(* Logix 5000 project; controller TFF vendor 1 type 14 code 107 rev 34.11; software revision 34.03; part 24 of 36 *)
(* tags used below, declared in another part *)
   Address : DINT;   // Temp Address
   Address2 : DINT;   // Temp Address
   Index : DINT;   // Index
   ONS_PID02 : BOOL;
   PCV001_PID_Settings : INT;
   AnalogOutput : AnalogOutput[25];   // Analog Output Array
   AnalogPoint : AnalogInput[50];   // Analog Input Array
   ControlLoop : ControlLoop[20];   // Control Loop Array
   ControlLoop_FeedPump : ALIAS FOR ControlLoop[1];   // Feed Pump Control Loop
   ControlLoop_PCV001 : ALIAS FOR ControlLoop[3];   // PCV001 Control Loop
   ControlLoop_PCV001_5ms : ALIAS FOR ControlLoop[4];   // PCV001 Control Loop
   ControlLoop_PCV001_CV : REAL;   // Control Value
   ControlLoop_PCV001_RAMP_OUT : REAL;   // Ramp Output
   ControlLoop_PCV101 : ALIAS FOR ControlLoop[5];   // PCV101 Control Loop
   ControlLoop_PCV101_5ms : ALIAS FOR ControlLoop[6];   // PCV101 Control Loop
   ControlLoop_PCV101_RAMP_OUT : REAL;   // Ramp Output
   PCV001_Control : PCV_Control;   // PCV001 Control UDT
   PCV101 : ALIAS FOR AnalogPoint[4];   // Filtrate Pressure Control Valve Position
   PCV101_Control : PCV_Control;   // PCV101 Control UDT
   PumpRunStatus : DINT;   // Pumps Run Status (1 = At least one pump running , 0 = no pump running)
   SysControl : SysControl;   // General system status and command
(* Process, continued *)

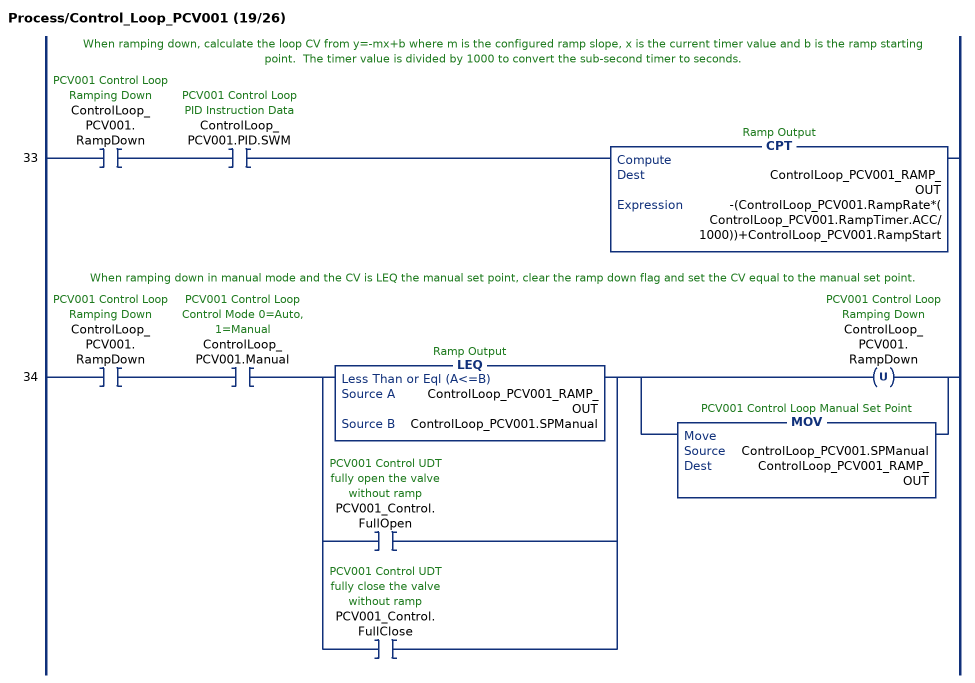
   [picture p213: Process/Control_Loop_PCV001 rungs 33-34]
   // When ramping down, calculate the loop CV from y=-mx+b where m is the configured ramp slope, x is the current timer value and b is the ramp starting point.  The timer value is divided by 1000 to convert the sub-second timer to seconds.
   33: XIC(ControlLoop_PCV001.RampDown)XIC(ControlLoop_PCV001.PID.SWM)CPT(ControlLoop_PCV001_RAMP_OUT,-(ControlLoop_PCV001.RampRate*(ControlLoop_PCV001.RampTimer.ACC/1000))+ControlLoop_PCV001.RampStart);
   // When ramping down in manual mode and the CV is LEQ the manual set point, clear the ramp down flag and set the CV equal to the manual set point.
   34: XIC(ControlLoop_PCV001.RampDown)XIC(ControlLoop_PCV001.Manual)[LEQ(ControlLoop_PCV001_RAMP_OUT,ControlLoop_PCV001.SPManual) ,XIC(PCV001_Control.FullOpen) ,XIC(PCV001_Control.FullClose) ][OTU(ControlLoop_PCV001.RampDown) ,MOV(ControlLoop_PCV001.SPManual,ControlLoop_PCV001_RAMP_OUT) ];
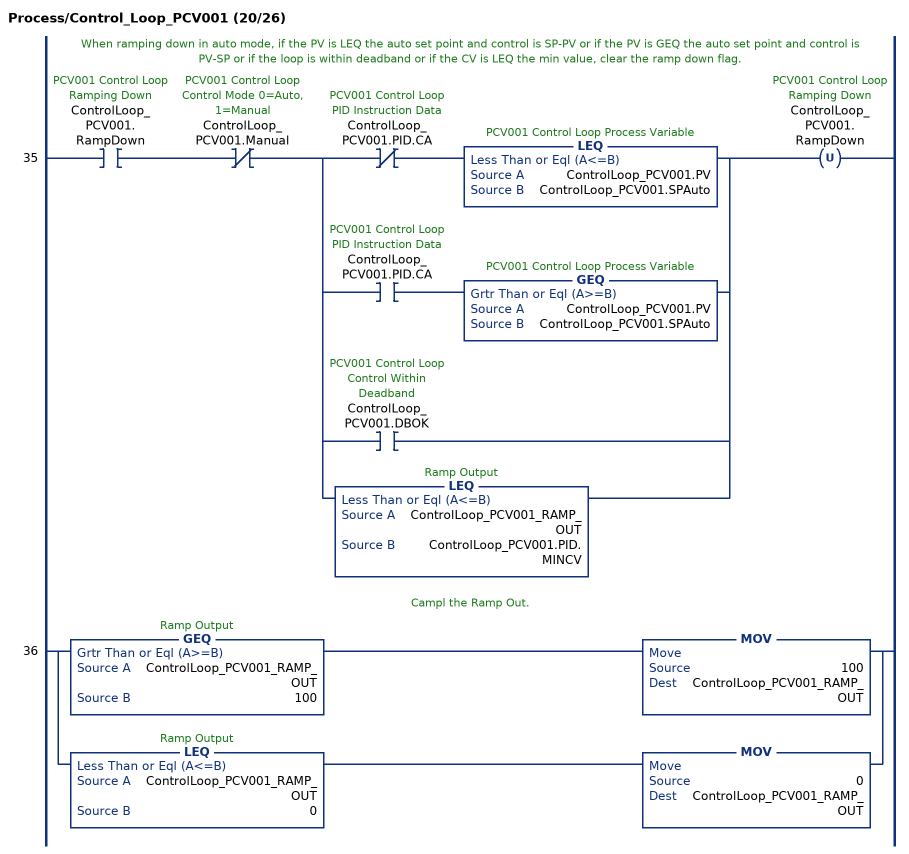
   // When ramping down in auto mode, if the PV is LEQ the auto set point and control is SP-PV or if the PV is GEQ the auto set point and control is PV-SP or if the loop is within deadband or if the CV is LEQ the min value, clear the ramp down flag.
   35: XIC(ControlLoop_PCV001.RampDown)XIO(ControlLoop_PCV001.Manual)[XIO(ControlLoop_PCV001.PID.CA) LEQ(ControlLoop_PCV001.PV,ControlLoop_PCV001.SPAuto) ,XIC(ControlLoop_PCV001.PID.CA) GEQ(ControlLoop_PCV001.PV,ControlLoop_PCV001.SPAuto) ,XIC(ControlLoop_PCV001.DBOK) ,LEQ(ControlLoop_PCV001_RAMP_OUT,ControlLoop_PCV001.PID.MINCV) ]OTU(ControlLoop_PCV001.RampDown);
   // Campl the Ramp Out.
   36: [GEQ(ControlLoop_PCV001_RAMP_OUT,100) MOV(100,ControlLoop_PCV001_RAMP_OUT) ,LEQ(ControlLoop_PCV001_RAMP_OUT,0) MOV(0,ControlLoop_PCV001_RAMP_OUT) ];
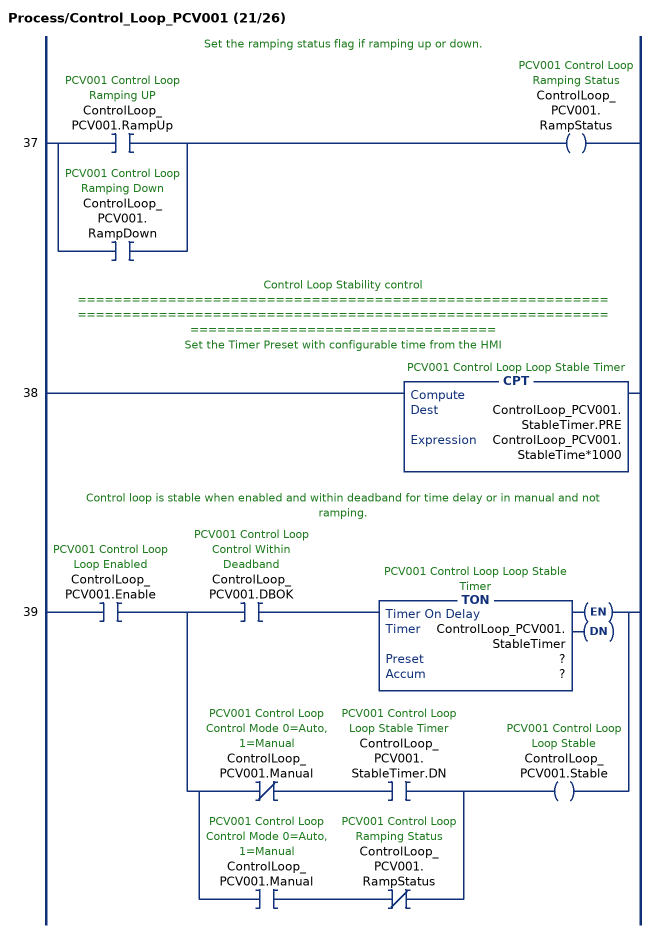
   // Set the ramping status flag if ramping up or down.
   37: [XIC(ControlLoop_PCV001.RampUp) ,XIC(ControlLoop_PCV001.RampDown) ]OTE(ControlLoop_PCV001.RampStatus);
   // Control Loop Stability control
   // ========================================================================================================================================================
   // Set the Timer Preset with configurable time from the HMI
   38: CPT(ControlLoop_PCV001.StableTimer.PRE,ControlLoop_PCV001.StableTime*1000);
   // Control loop is stable when enabled and within deadband for time delay or in manual and not ramping.
   39: XIC(ControlLoop_PCV001.Enable)[XIC(ControlLoop_PCV001.DBOK) TON(ControlLoop_PCV001.StableTimer,?,?) ,[XIO(ControlLoop_PCV001.Manual) XIC(ControlLoop_PCV001.StableTimer.DN) ,XIC(ControlLoop_PCV001.Manual) XIO(ControlLoop_PCV001.RampStatus) ] OTE(ControlLoop_PCV001.Stable) ];
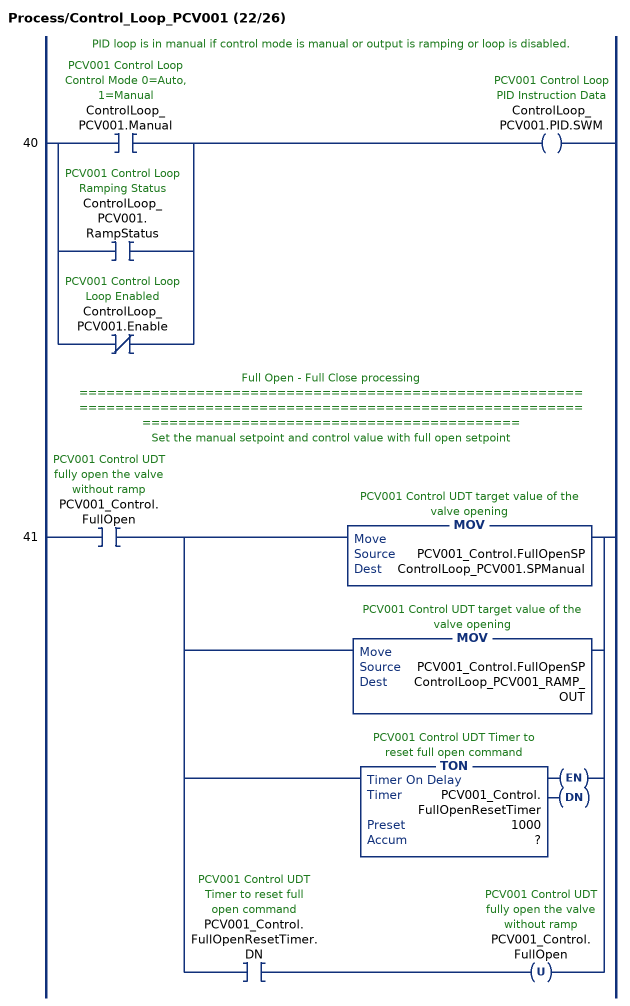
   // PID loop is in manual if control mode is manual or output is ramping or loop is disabled.
   40: [XIC(ControlLoop_PCV001.Manual) ,XIC(ControlLoop_PCV001.RampStatus) ,XIO(ControlLoop_PCV001.Enable) ]OTE(ControlLoop_PCV001.PID.SWM);
   // Full Open - Full Close processing
   // ==========================================================================================================================================================
   // Set the manual setpoint and control value with full open setpoint
   41: XIC(PCV001_Control.FullOpen)[MOV(PCV001_Control.FullOpenSP,ControlLoop_PCV001.SPManual) ,MOV(PCV001_Control.FullOpenSP,ControlLoop_PCV001_RAMP_OUT) ,TON(PCV001_Control.FullOpenResetTimer,?,?) ,XIC(PCV001_Control.FullOpenResetTimer.DN) OTU(PCV001_Control.FullOpen) ];
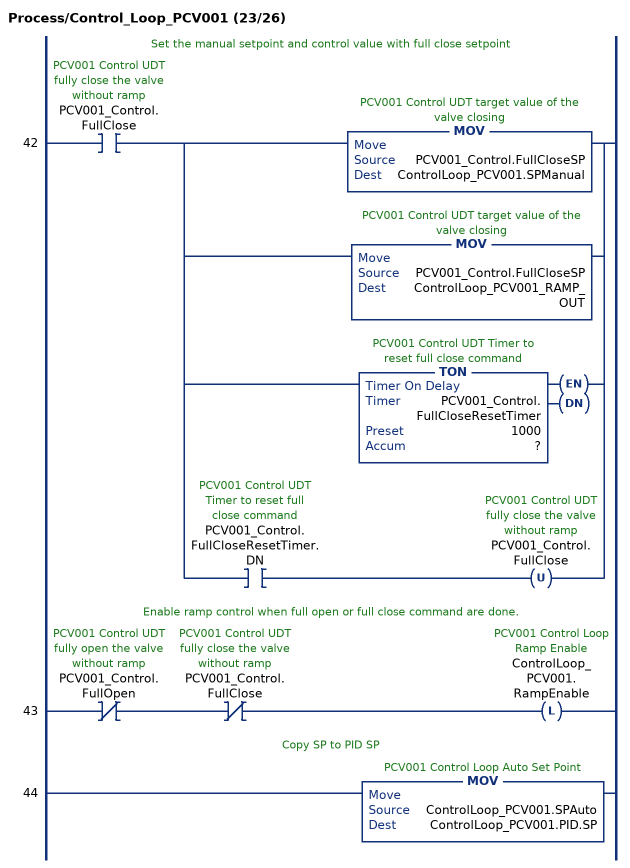
   // Set the manual setpoint and control value with full close setpoint
   42: XIC(PCV001_Control.FullClose)[MOV(PCV001_Control.FullCloseSP,ControlLoop_PCV001.SPManual) ,MOV(PCV001_Control.FullCloseSP,ControlLoop_PCV001_RAMP_OUT) ,TON(PCV001_Control.FullCloseResetTimer,?,?) ,XIC(PCV001_Control.FullCloseResetTimer.DN) OTU(PCV001_Control.FullClose) ];
   // Enable ramp control when full open or full close command are done.
   43: XIO(PCV001_Control.FullOpen)XIO(PCV001_Control.FullClose)OTL(ControlLoop_PCV001.RampEnable);
   // Copy SP to PID SP
   44: MOV(ControlLoop_PCV001.SPAuto,ControlLoop_PCV001.PID.SP);
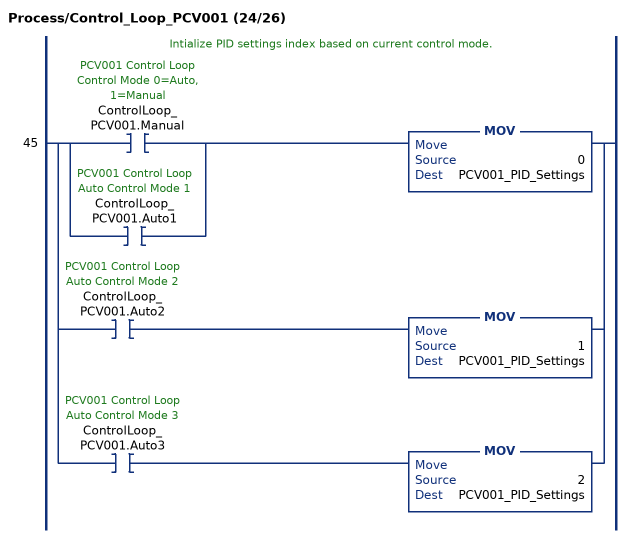
   // Intialize PID settings index based on current control mode.
   45: [[XIC(ControlLoop_PCV001.Manual) ,XIC(ControlLoop_PCV001.Auto1) ] MOV(0,PCV001_PID_Settings) ,XIC(ControlLoop_PCV001.Auto2) MOV(1,PCV001_PID_Settings) ,XIC(ControlLoop_PCV001.Auto3) MOV(2,PCV001_PID_Settings) ];
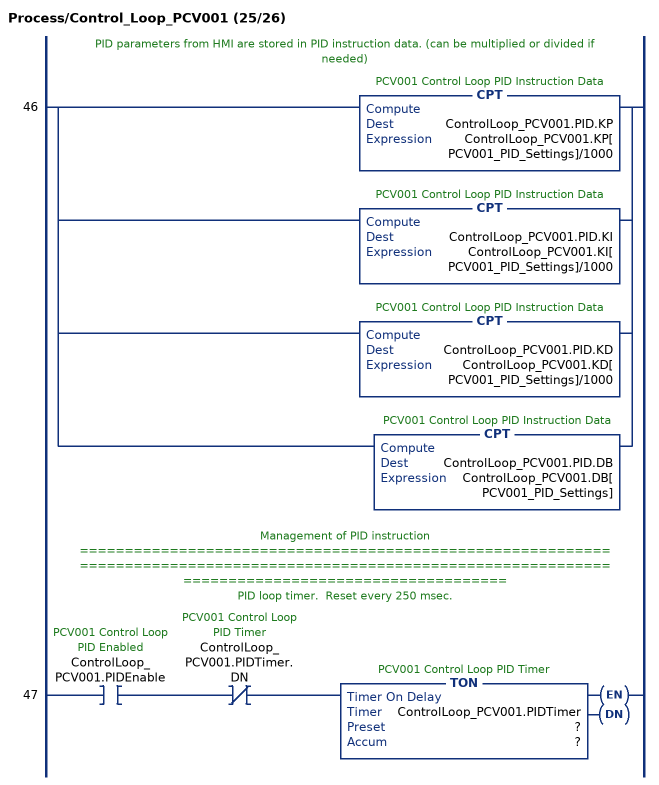
   // PID parameters from HMI are stored in PID instruction data. (can be multiplied or divided if needed)
   46: [CPT(ControlLoop_PCV001.PID.KP,ControlLoop_PCV001.KP[PCV001_PID_Settings]/1000) ,CPT(ControlLoop_PCV001.PID.KI,ControlLoop_PCV001.KI[PCV001_PID_Settings]/1000) ,CPT(ControlLoop_PCV001.PID.KD,ControlLoop_PCV001.KD[PCV001_PID_Settings]/1000) ,CPT(ControlLoop_PCV001.PID.DB,ControlLoop_PCV001.DB[PCV001_PID_Settings]) ];
   // Management of PID instruction
   // ==========================================================================================================================================================
   // PID loop timer.  Reset every 250 msec.
   47: XIC(ControlLoop_PCV001.PIDEnable)XIO(ControlLoop_PCV001.PIDTimer.DN)TON(ControlLoop_PCV001.PIDTimer,?,?);
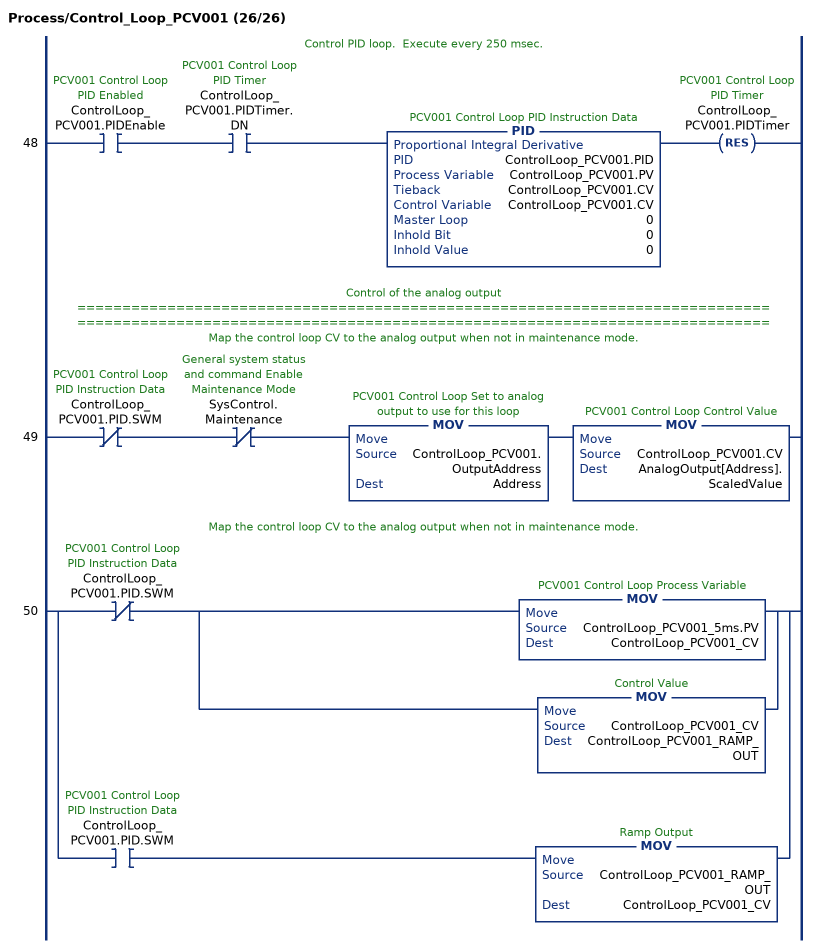
   // Control PID loop.  Execute every 250 msec.
   48: XIC(ControlLoop_PCV001.PIDEnable)XIC(ControlLoop_PCV001.PIDTimer.DN)PID(ControlLoop_PCV001.PID,ControlLoop_PCV001.PV,ControlLoop_PCV001.CV,ControlLoop_PCV001.CV,0,0,0)RES(ControlLoop_PCV001.PIDTimer);
   // Control of the analog output
   // ==========================================================================================================================================================
   // Map the control loop CV to the analog output when not in maintenance mode.
   49: XIO(ControlLoop_PCV001.PID.SWM)XIO(SysControl.Maintenance)MOV(ControlLoop_PCV001.OutputAddress,Address)MOV(ControlLoop_PCV001.CV,AnalogOutput[Address].ScaledValue);
   // Map the control loop CV to the analog output when not in maintenance mode.
   50: [XIO(ControlLoop_PCV001.PID.SWM) [MOV(ControlLoop_PCV001_5ms.PV,ControlLoop_PCV001_CV) ,MOV(ControlLoop_PCV001_CV,ControlLoop_PCV001_RAMP_OUT) ] ,XIC(ControlLoop_PCV001.PID.SWM) MOV(ControlLoop_PCV001_RAMP_OUT,ControlLoop_PCV001_CV) ];
END_ROUTINE

ROUTINE Control_Loop_PCV101   (* ladder *)
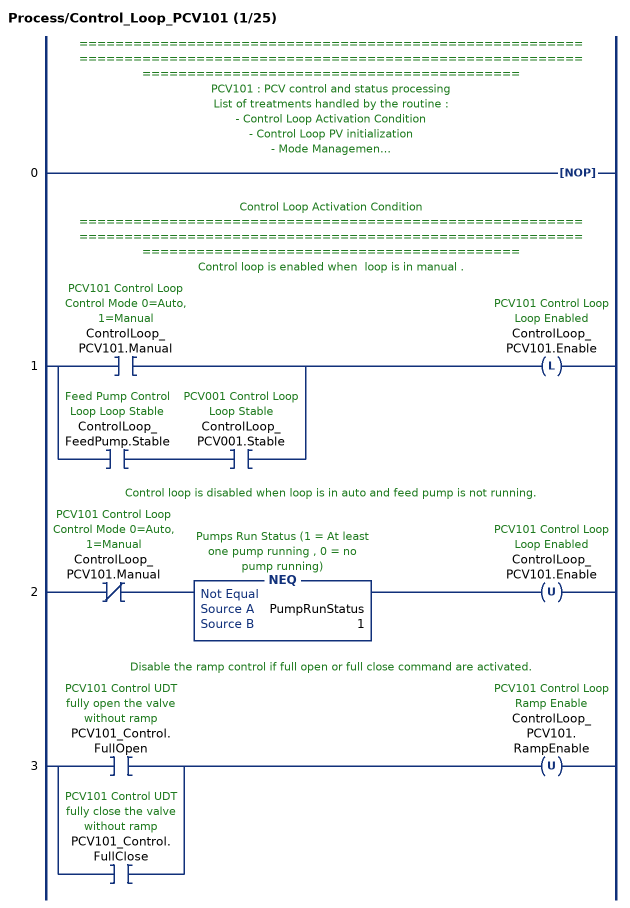
   // ==========================================================================================================================================================
   //                                                  PCV101 : PCV control and status processing
   //                                                     List of treatments handled by the routine :
   //                                                          - Control Loop Activation Condition
   //                                                  - Control Loop PV initialization
   //                                                - Mode Management
   //                                                        - Control Loop Setpoint management
   //                                                        - Control Loop deadband calculation
   //                                                          - Management of ramping control
   //                                                          - Control Loop Stability control
   //                                                          - Full Open - Full Close processing
   //                                                          - Management of PID instruction
   //                                                          - Control of the analog output
   //                                                     -----------------------------------------------------------------------------------------------------------------------------------------------------
   //                                                     History
   //                                                          2019-SEP-26 - Actemium - B. Roch - Initial version for Candidate Release 3.00.00.00.c
   //      2019-OCT-25 - Actemium - B. Roch - Modification for Candidate Release 3.00.00.00.d
   //                                                    - delete the mode change action on default state
   //     2020-SEP-14 - Merck - Q. Spindler - Modifications for Candidate Release 3.00.00.01.a
   //                                                        - on rung 16, disable DBOK if control loop is not enabled or in manual
   // 	   2021-APR-19 - DAVIDSON- Ch. ARBOGAST - Modifications for Candidate Release 3.01.00.00.a
   // 	- on rung 4, line 1, replace "ControlLoop[5].Manual OR ControlLoop[5].Auto1" by
   // 			 "NOT ControlLoop[5].Auto2 AND NOT ControlLoop[5].Auto3"
   // ==========================================================================================================================================================
   0: NOP();
   // Control Loop Activation Condition
   // ==========================================================================================================================================================
   // Control loop is enabled when  loop is in manual .
   1: [XIC(ControlLoop_PCV101.Manual) ,XIC(ControlLoop_FeedPump.Stable) XIC(ControlLoop_PCV001.Stable) ]OTL(ControlLoop_PCV101.Enable);
   // Control loop is disabled when loop is in auto and feed pump is not running.
   2: XIO(ControlLoop_PCV101.Manual)NEQ(PumpRunStatus,1)OTU(ControlLoop_PCV101.Enable);
   // Disable the ramp control if full open or full close command are activated.
   3: [XIC(PCV101_Control.FullOpen) ,XIC(PCV101_Control.FullClose) ]OTU(ControlLoop_PCV101.RampEnable);
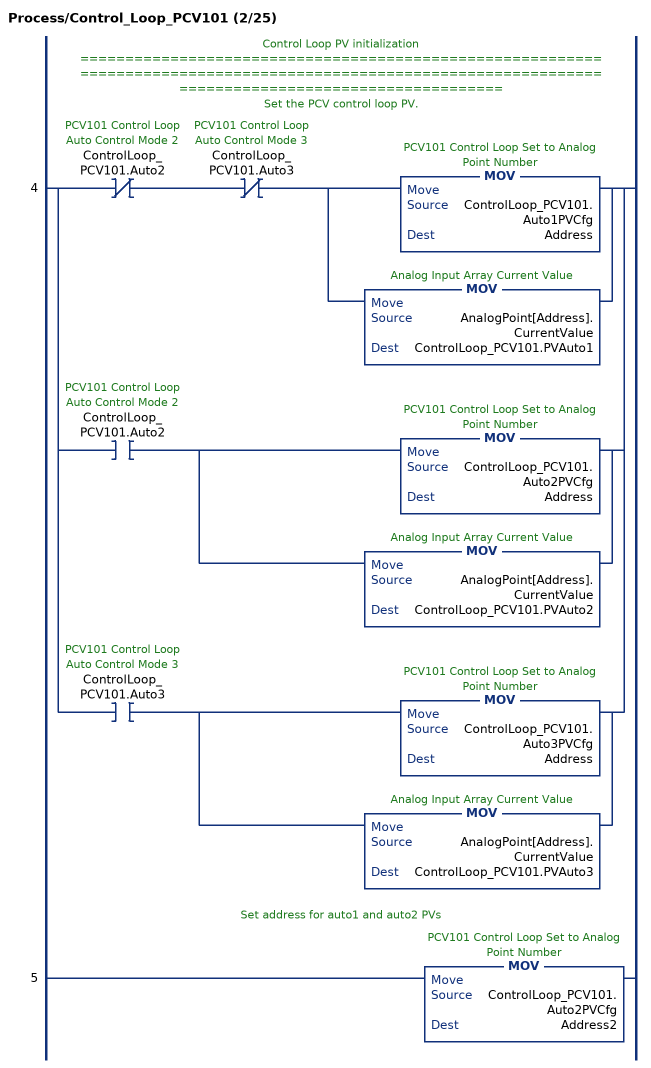
   // Control Loop PV initialization
   // ========================================================================================================================================================
   // Set the PCV control loop PV.
   4: [[XIO(ControlLoop_PCV101.Auto2) XIO(ControlLoop_PCV101.Auto3) [MOV(ControlLoop_PCV101.Auto1PVCfg,Address) ,MOV(AnalogPoint[Address].CurrentValue,ControlLoop_PCV101.PVAuto1) ] ,XIC(ControlLoop_PCV101.Auto2) [MOV(ControlLoop_PCV101.Auto2PVCfg,Address) ,MOV(AnalogPoint[Address].CurrentValue,ControlLoop_PCV101.PVAuto2) ] ] ,XIC(ControlLoop_PCV101.Auto3) [MOV(ControlLoop_PCV101.Auto3PVCfg,Address) ,MOV(AnalogPoint[Address].CurrentValue,ControlLoop_PCV101.PVAuto3) ] ];
   // Set address for auto1 and auto2 PVs
   5: MOV(ControlLoop_PCV101.Auto2PVCfg,Address2);
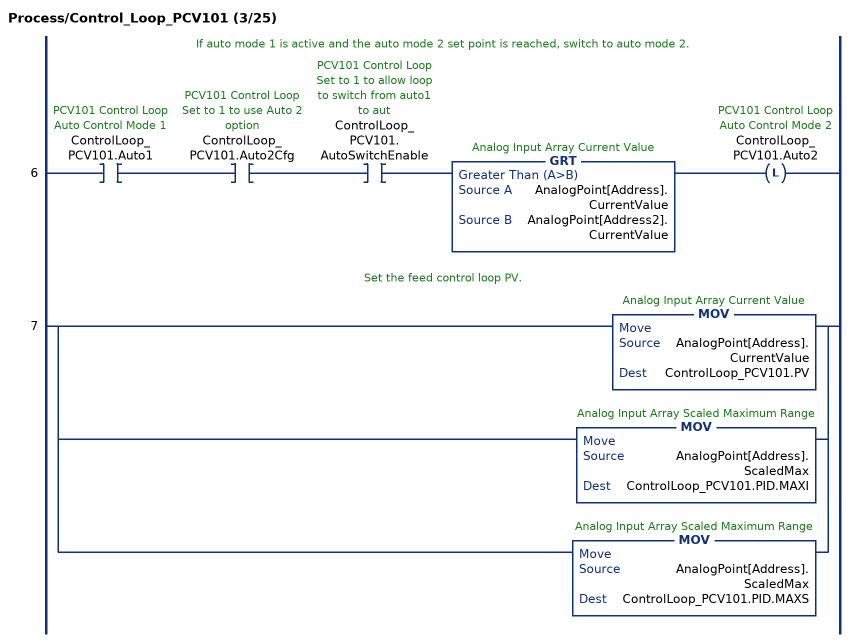
   // If auto mode 1 is active and the auto mode 2 set point is reached, switch to auto mode 2.
   6: XIC(ControlLoop_PCV101.Auto1)XIC(ControlLoop_PCV101.Auto2Cfg)XIC(ControlLoop_PCV101.AutoSwitchEnable)GRT(AnalogPoint[Address].CurrentValue,AnalogPoint[Address2].CurrentValue)OTL(ControlLoop_PCV101.Auto2);
   // Set the feed control loop PV.
   7: [MOV(AnalogPoint[Address].CurrentValue,ControlLoop_PCV101.PV) ,MOV(AnalogPoint[Address].ScaledMax,ControlLoop_PCV101.PID.MAXI) ,MOV(AnalogPoint[Address].ScaledMax,ControlLoop_PCV101.PID.MAXS) ];
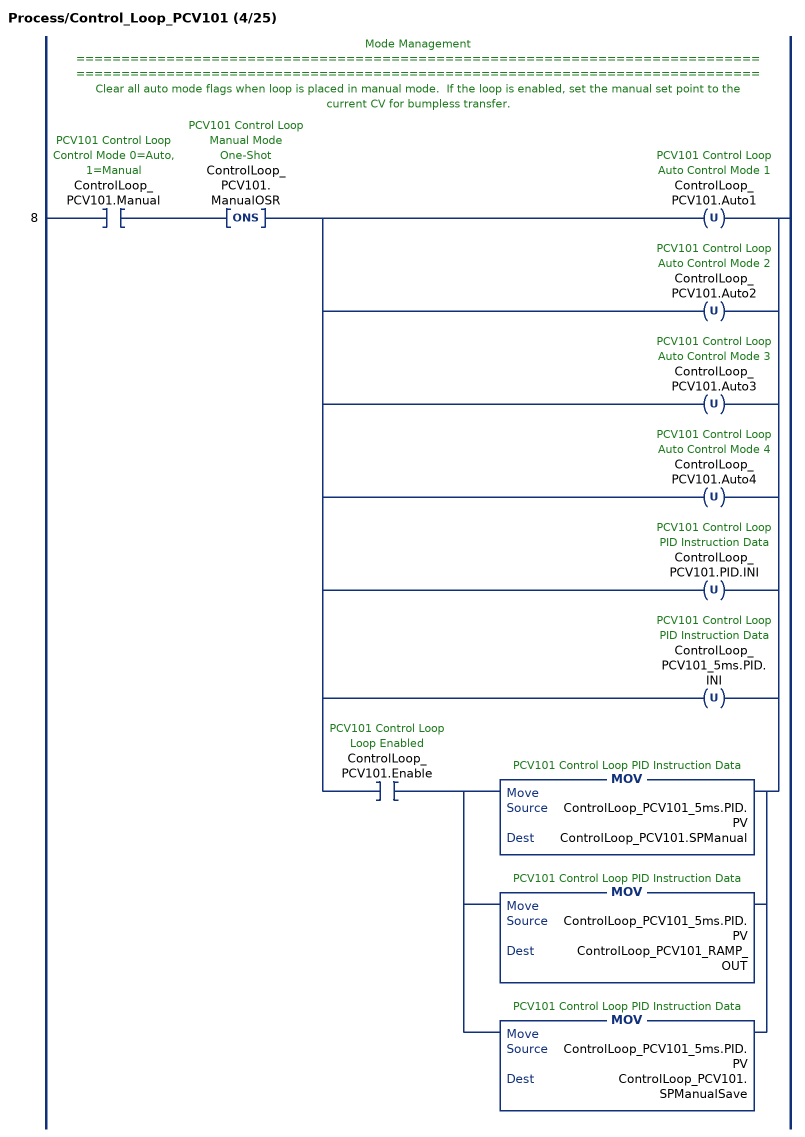
   // Mode Management
   // ========================================================================================================================================================
   // Clear all auto mode flags when loop is placed in manual mode.  If the loop is enabled, set the manual set point to the current CV for bumpless transfer.
   8: XIC(ControlLoop_PCV101.Manual)ONS(ControlLoop_PCV101.ManualOSR)[OTU(ControlLoop_PCV101.Auto1) ,OTU(ControlLoop_PCV101.Auto2) ,OTU(ControlLoop_PCV101.Auto3) ,OTU(ControlLoop_PCV101.Auto4) ,OTU(ControlLoop_PCV101.PID.INI) ,OTU(ControlLoop_PCV101_5ms.PID.INI) ,XIC(ControlLoop_PCV101.Enable) [MOV(ControlLoop_PCV101_5ms.PID.PV,ControlLoop_PCV101.SPManual) ,MOV(ControlLoop_PCV101_5ms.PID.PV,ControlLoop_PCV101_RAMP_OUT) ,MOV(ControlLoop_PCV101_5ms.PID.PV,ControlLoop_PCV101.SPManualSave) ] ];
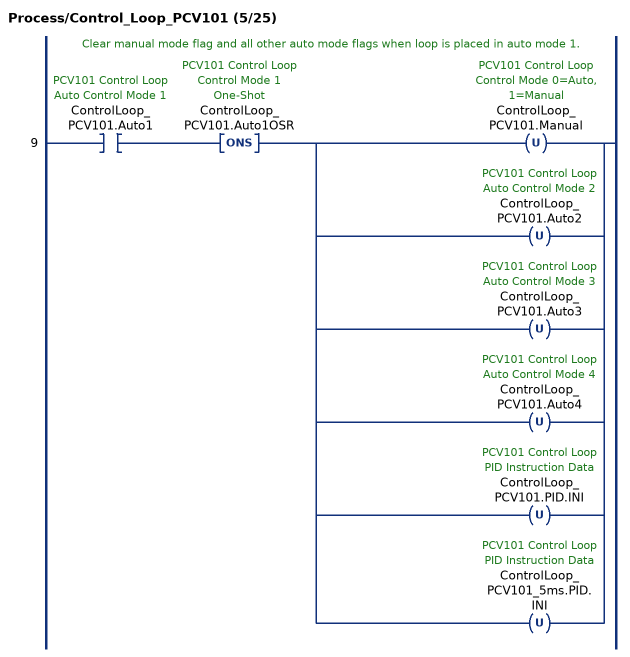
   // Clear manual mode flag and all other auto mode flags when loop is placed in auto mode 1.
   9: XIC(ControlLoop_PCV101.Auto1)ONS(ControlLoop_PCV101.Auto1OSR)[OTU(ControlLoop_PCV101.Manual) ,OTU(ControlLoop_PCV101.Auto2) ,OTU(ControlLoop_PCV101.Auto3) ,OTU(ControlLoop_PCV101.Auto4) ,OTU(ControlLoop_PCV101.PID.INI) ,OTU(ControlLoop_PCV101_5ms.PID.INI) ];
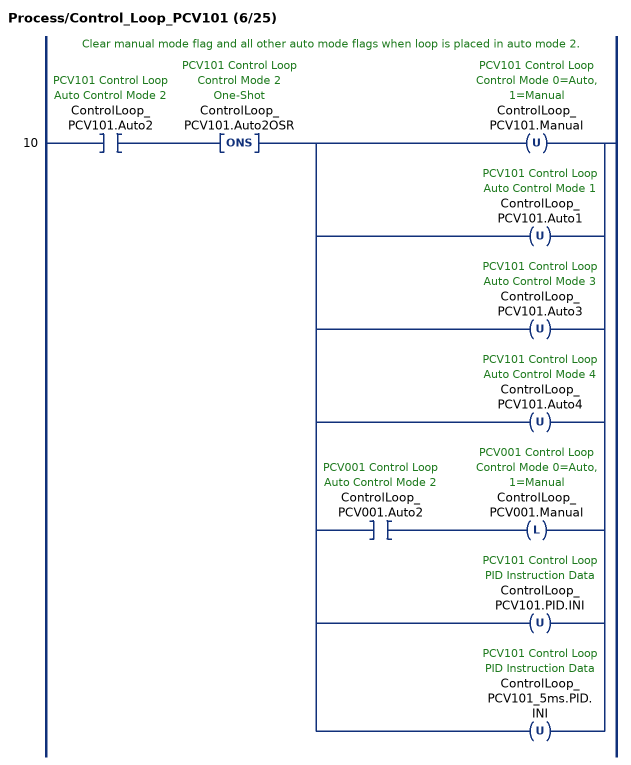
   // Clear manual mode flag and all other auto mode flags when loop is placed in auto mode 2.
   10: XIC(ControlLoop_PCV101.Auto2)ONS(ControlLoop_PCV101.Auto2OSR)[OTU(ControlLoop_PCV101.Manual) ,OTU(ControlLoop_PCV101.Auto1) ,OTU(ControlLoop_PCV101.Auto3) ,OTU(ControlLoop_PCV101.Auto4) ,XIC(ControlLoop_PCV001.Auto2) OTL(ControlLoop_PCV001.Manual) ,OTU(ControlLoop_PCV101.PID.INI) ,OTU(ControlLoop_PCV101_5ms.PID.INI) ];
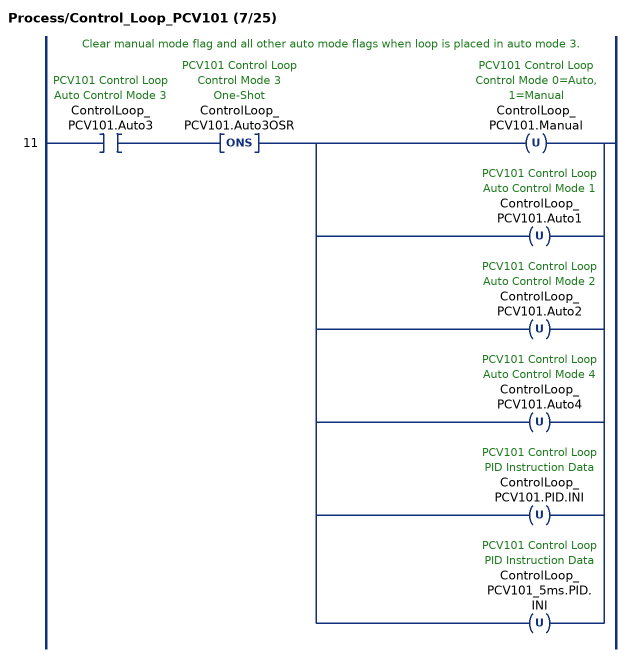
   // Clear manual mode flag and all other auto mode flags when loop is placed in auto mode 3.
   11: XIC(ControlLoop_PCV101.Auto3)ONS(ControlLoop_PCV101.Auto3OSR)[OTU(ControlLoop_PCV101.Manual) ,OTU(ControlLoop_PCV101.Auto1) ,OTU(ControlLoop_PCV101.Auto2) ,OTU(ControlLoop_PCV101.Auto4) ,OTU(ControlLoop_PCV101.PID.INI) ,OTU(ControlLoop_PCV101_5ms.PID.INI) ];
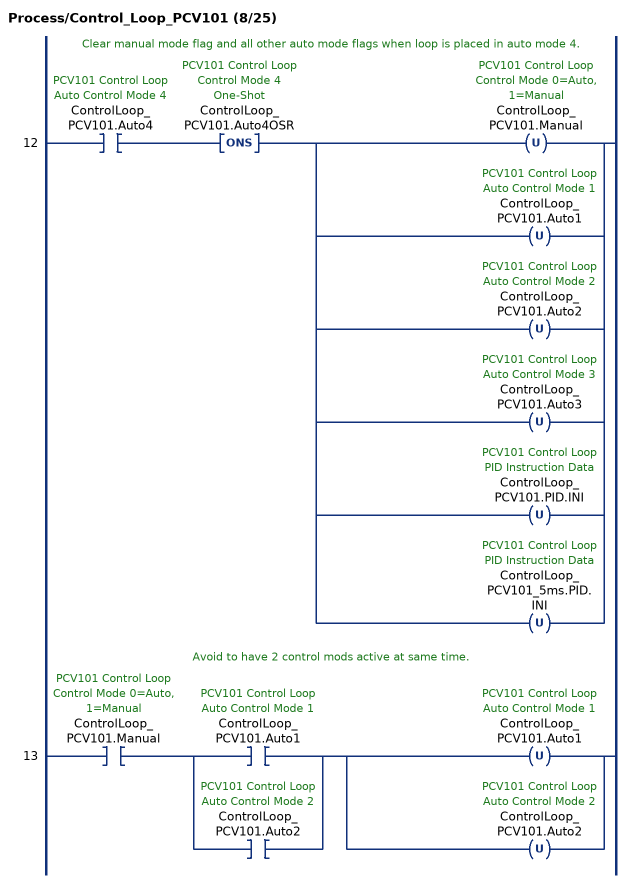
   // Clear manual mode flag and all other auto mode flags when loop is placed in auto mode 4.
   12: XIC(ControlLoop_PCV101.Auto4)ONS(ControlLoop_PCV101.Auto4OSR)[OTU(ControlLoop_PCV101.Manual) ,OTU(ControlLoop_PCV101.Auto1) ,OTU(ControlLoop_PCV101.Auto2) ,OTU(ControlLoop_PCV101.Auto3) ,OTU(ControlLoop_PCV101.PID.INI) ,OTU(ControlLoop_PCV101_5ms.PID.INI) ];
   // Avoid to have 2 control mods active at same time.
   13: XIC(ControlLoop_PCV101.Manual)[XIC(ControlLoop_PCV101.Auto1) ,XIC(ControlLoop_PCV101.Auto2) ][OTU(ControlLoop_PCV101.Auto1) ,OTU(ControlLoop_PCV101.Auto2) ];
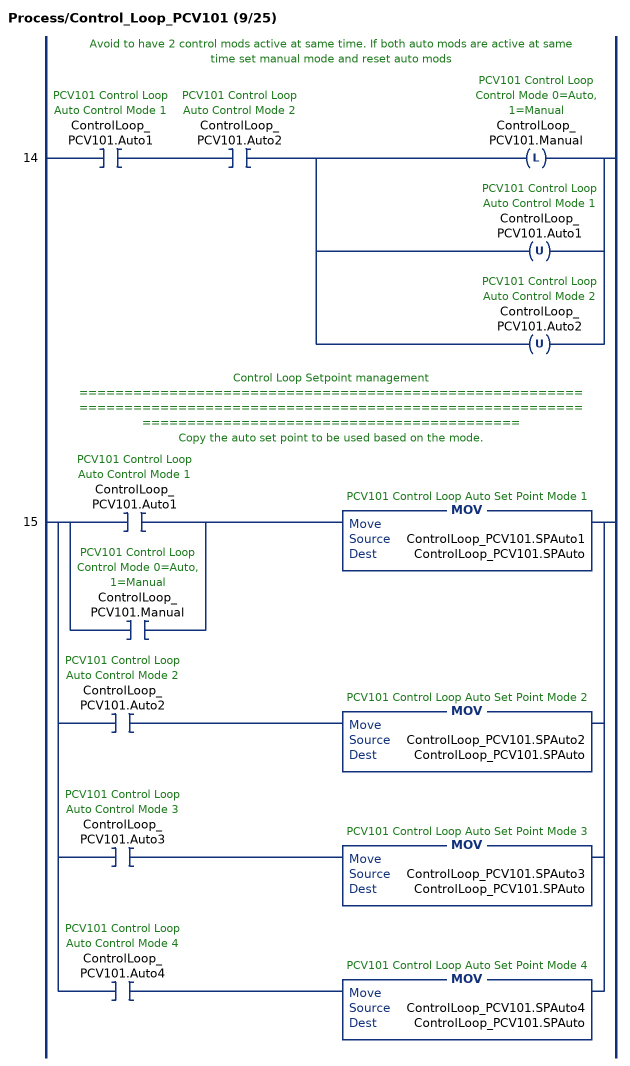
   // Avoid to have 2 control mods active at same time. If both auto mods are active at same time set manual mode and reset auto mods
   14: XIC(ControlLoop_PCV101.Auto1)XIC(ControlLoop_PCV101.Auto2)[OTL(ControlLoop_PCV101.Manual) ,OTU(ControlLoop_PCV101.Auto1) ,OTU(ControlLoop_PCV101.Auto2) ];
   // Control Loop Setpoint management
   // ==========================================================================================================================================================
   // Copy the auto set point to be used based on the mode.
   15: [[XIC(ControlLoop_PCV101.Auto1) ,XIC(ControlLoop_PCV101.Manual) ] MOV(ControlLoop_PCV101.SPAuto1,ControlLoop_PCV101.SPAuto) ,XIC(ControlLoop_PCV101.Auto2) MOV(ControlLoop_PCV101.SPAuto2,ControlLoop_PCV101.SPAuto) ,XIC(ControlLoop_PCV101.Auto3) MOV(ControlLoop_PCV101.SPAuto3,ControlLoop_PCV101.SPAuto) ,XIC(ControlLoop_PCV101.Auto4) MOV(ControlLoop_PCV101.SPAuto4,ControlLoop_PCV101.SPAuto) ];
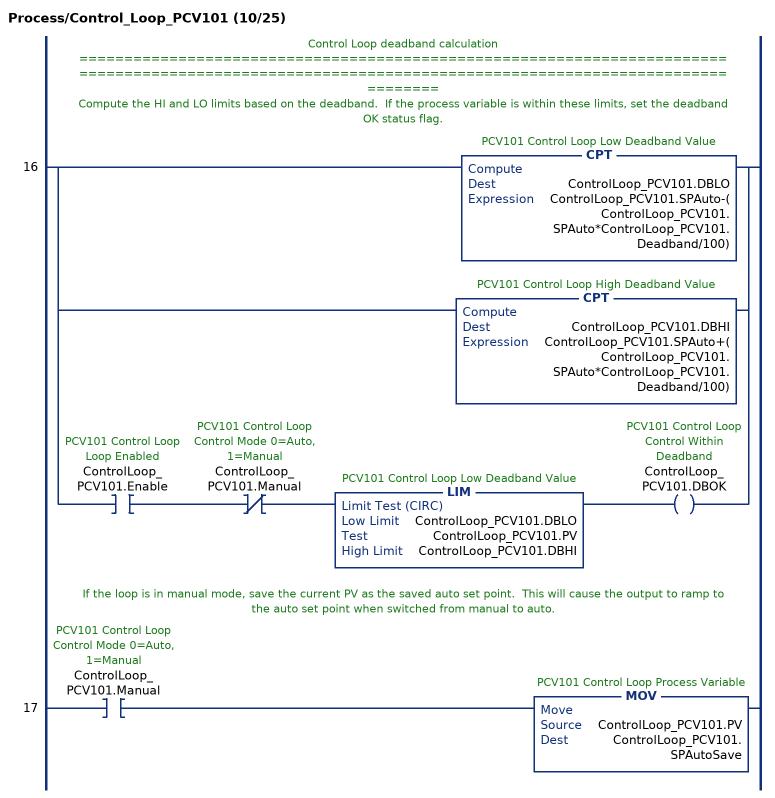
   // Control Loop deadband calculation
   // ========================================================================================================================================================
   // Compute the HI and LO limits based on the deadband.  If the process variable is within these limits, set the deadband OK status flag.
   16: [CPT(ControlLoop_PCV101.DBLO,ControlLoop_PCV101.SPAuto-(ControlLoop_PCV101.SPAuto*ControlLoop_PCV101.Deadband/100)) ,CPT(ControlLoop_PCV101.DBHI,ControlLoop_PCV101.SPAuto+(ControlLoop_PCV101.SPAuto*ControlLoop_PCV101.Deadband/100)) ,XIC(ControlLoop_PCV101.Enable) XIO(ControlLoop_PCV101.Manual) LIM(ControlLoop_PCV101.DBLO,ControlLoop_PCV101.PV,ControlLoop_PCV101.DBHI) OTE(ControlLoop_PCV101.DBOK) ];
   // If the loop is in manual mode, save the current PV as the saved auto set point.  This will cause the output to ramp to the auto set point when switched from manual to auto.
   17: XIC(ControlLoop_PCV101.Manual)MOV(ControlLoop_PCV101.PV,ControlLoop_PCV101.SPAutoSave);
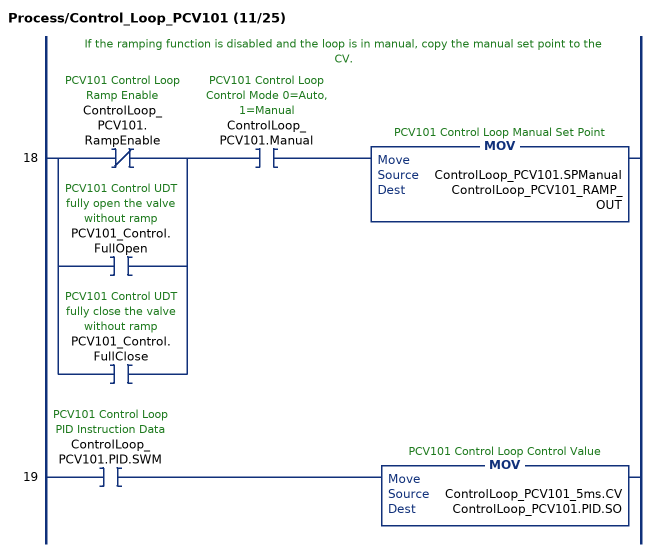
   // If the ramping function is disabled and the loop is in manual, copy the manual set point to the CV.
   18: [XIO(ControlLoop_PCV101.RampEnable) ,XIC(PCV101_Control.FullOpen) ,XIC(PCV101_Control.FullClose) ]XIC(ControlLoop_PCV101.Manual)MOV(ControlLoop_PCV101.SPManual,ControlLoop_PCV101_RAMP_OUT);
   19: XIC(ControlLoop_PCV101.PID.SWM)MOV(ControlLoop_PCV101_5ms.CV,ControlLoop_PCV101.PID.SO);
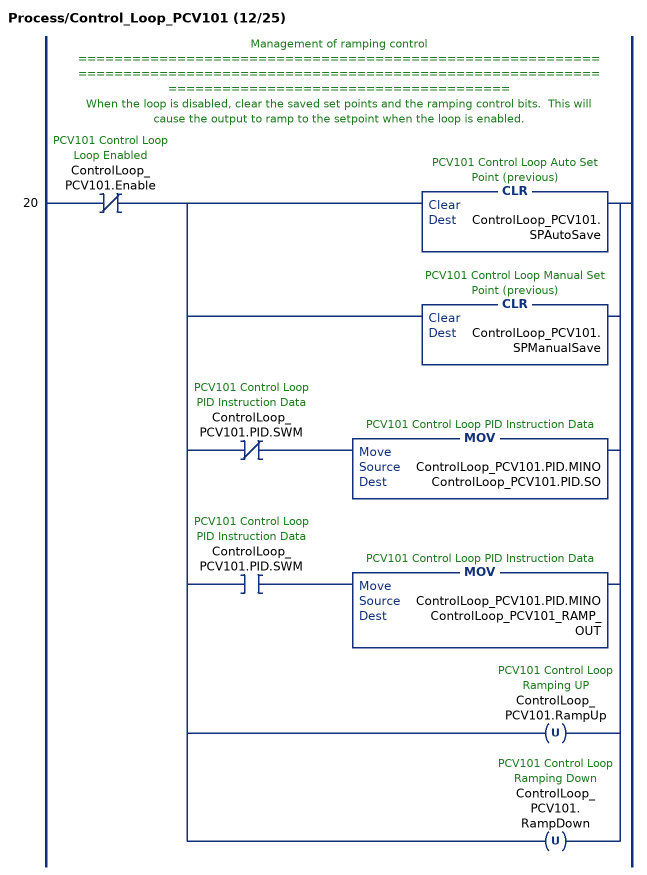
   // Management of ramping control
   // ==========================================================================================================================================================
   // When the loop is disabled, clear the saved set points and the ramping control bits.  This will cause the output to ramp to the setpoint when the loop is enabled.
   20: XIO(ControlLoop_PCV101.Enable)[CLR(ControlLoop_PCV101.SPAutoSave) ,CLR(ControlLoop_PCV101.SPManualSave) ,XIO(ControlLoop_PCV101.PID.SWM) MOV(ControlLoop_PCV101.PID.MINO,ControlLoop_PCV101.PID.SO) ,XIC(ControlLoop_PCV101.PID.SWM) MOV(ControlLoop_PCV101.PID.MINO,ControlLoop_PCV101_RAMP_OUT) ,OTU(ControlLoop_PCV101.RampUp) ,OTU(ControlLoop_PCV101.RampDown) ];
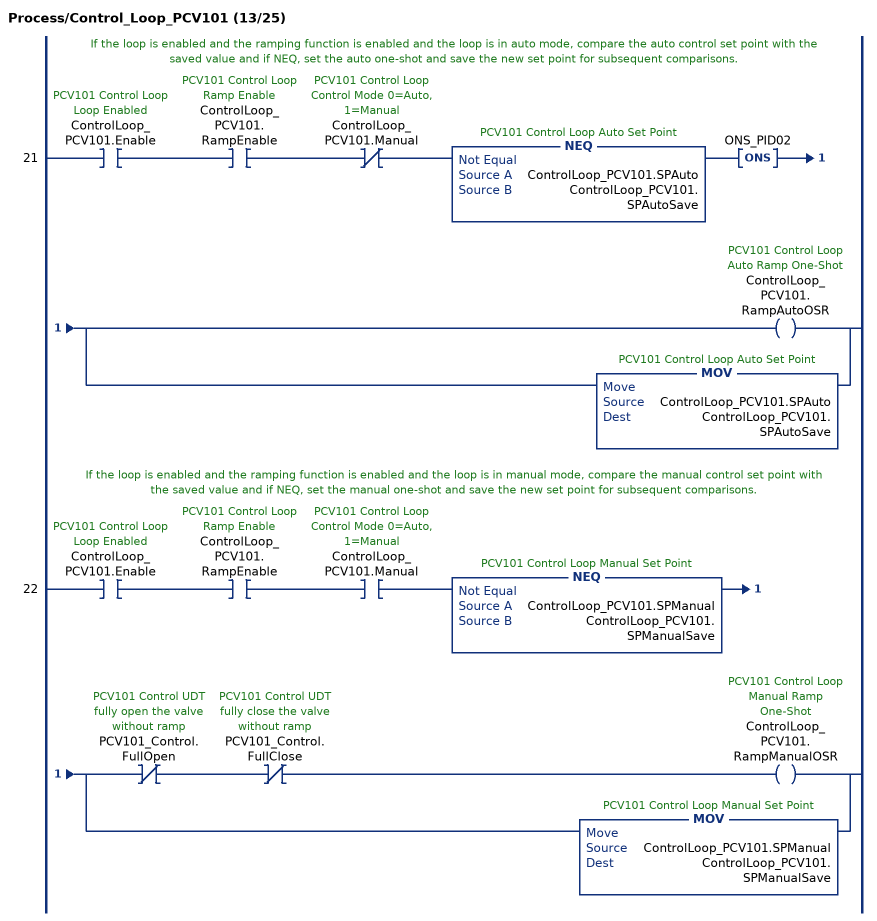
   // If the loop is enabled and the ramping function is enabled and the loop is in auto mode, compare the auto control set point with the saved value and if NEQ, set the auto one-shot and save the new set point for subsequent comparisons.
   21: XIC(ControlLoop_PCV101.Enable)XIC(ControlLoop_PCV101.RampEnable)XIO(ControlLoop_PCV101.Manual)NEQ(ControlLoop_PCV101.SPAuto,ControlLoop_PCV101.SPAutoSave)ONS(ONS_PID02)[OTE(ControlLoop_PCV101.RampAutoOSR) ,MOV(ControlLoop_PCV101.SPAuto,ControlLoop_PCV101.SPAutoSave) ];
   // If the loop is enabled and the ramping function is enabled and the loop is in manual mode, compare the manual control set point with the saved value and if NEQ, set the manual one-shot and save the new set point for subsequent comparisons.
   22: XIC(ControlLoop_PCV101.Enable)XIC(ControlLoop_PCV101.RampEnable)XIC(ControlLoop_PCV101.Manual)NEQ(ControlLoop_PCV101.SPManual,ControlLoop_PCV101.SPManualSave)[XIO(PCV101_Control.FullOpen) XIO(PCV101_Control.FullClose) OTE(ControlLoop_PCV101.RampManualOSR) ,MOV(ControlLoop_PCV101.SPManual,ControlLoop_PCV101.SPManualSave) ];
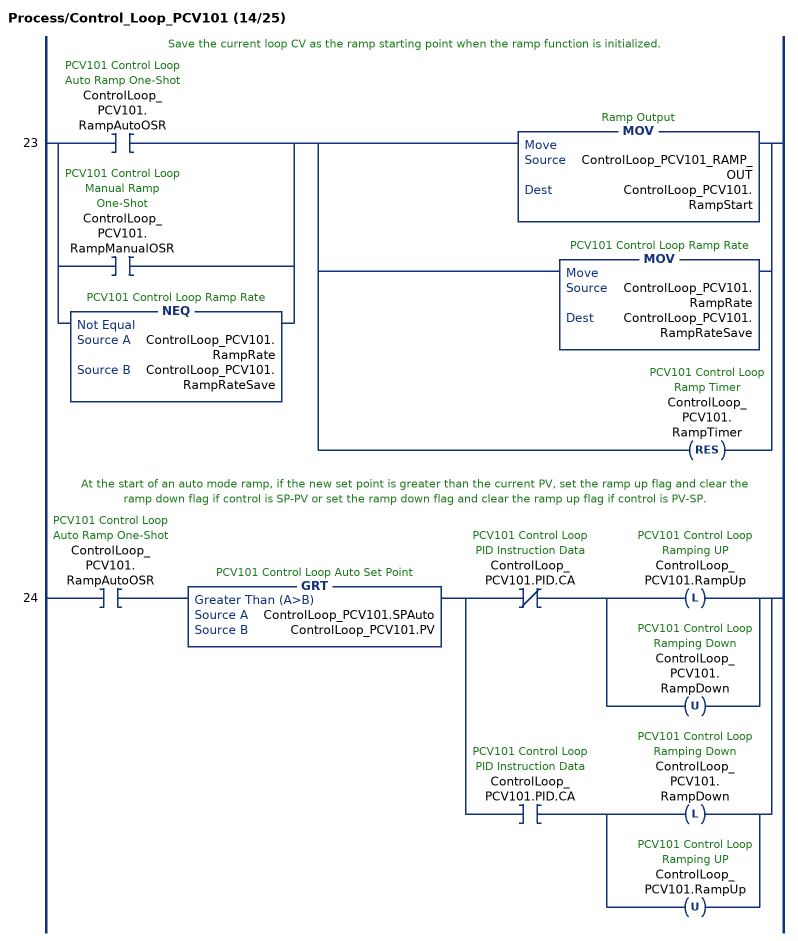
   // Save the current loop CV as the ramp starting point when the ramp function is initialized.
   23: [XIC(ControlLoop_PCV101.RampAutoOSR) ,XIC(ControlLoop_PCV101.RampManualOSR) ,NEQ(ControlLoop_PCV101.RampRate,ControlLoop_PCV101.RampRateSave) ][MOV(ControlLoop_PCV101_RAMP_OUT,ControlLoop_PCV101.RampStart) ,MOV(ControlLoop_PCV101.RampRate,ControlLoop_PCV101.RampRateSave) ,RES(ControlLoop_PCV101.RampTimer) ];
   // At the start of an auto mode ramp, if the new set point is greater than the current PV, set the ramp up flag and clear the ramp down flag if control is SP-PV or set the ramp down flag and clear the ramp up flag if control is PV-SP.
   24: XIC(ControlLoop_PCV101.RampAutoOSR)GRT(ControlLoop_PCV101.SPAuto,ControlLoop_PCV101.PV)[XIO(ControlLoop_PCV101.PID.CA) [OTL(ControlLoop_PCV101.RampUp) ,OTU(ControlLoop_PCV101.RampDown) ] ,XIC(ControlLoop_PCV101.PID.CA) [OTL(ControlLoop_PCV101.RampDown) ,OTU(ControlLoop_PCV101.RampUp) ] ];
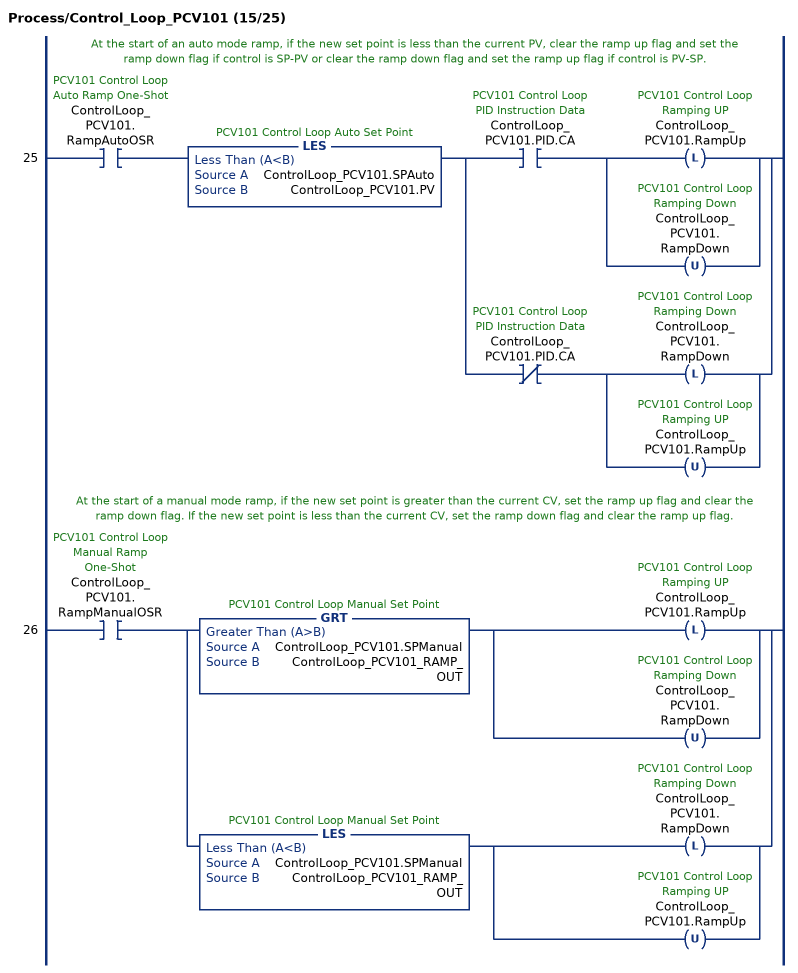
   // At the start of an auto mode ramp, if the new set point is less than the current PV, clear the ramp up flag and set the ramp down flag if control is SP-PV or clear the ramp down flag and set the ramp up flag if control is PV-SP.
   25: XIC(ControlLoop_PCV101.RampAutoOSR)LES(ControlLoop_PCV101.SPAuto,ControlLoop_PCV101.PV)[XIC(ControlLoop_PCV101.PID.CA) [OTL(ControlLoop_PCV101.RampUp) ,OTU(ControlLoop_PCV101.RampDown) ] ,XIO(ControlLoop_PCV101.PID.CA) [OTL(ControlLoop_PCV101.RampDown) ,OTU(ControlLoop_PCV101.RampUp) ] ];
   // At the start of a manual mode ramp, if the new set point is greater than the current CV, set the ramp up flag and clear the ramp down flag. If the new set point is less than the current CV, set the ramp down flag and clear the ramp up flag.
   26: XIC(ControlLoop_PCV101.RampManualOSR)[GRT(ControlLoop_PCV101.SPManual,ControlLoop_PCV101_RAMP_OUT) [OTL(ControlLoop_PCV101.RampUp) ,OTU(ControlLoop_PCV101.RampDown) ] ,LES(ControlLoop_PCV101.SPManual,ControlLoop_PCV101_RAMP_OUT) [OTL(ControlLoop_PCV101.RampDown) ,OTU(ControlLoop_PCV101.RampUp) ] ];
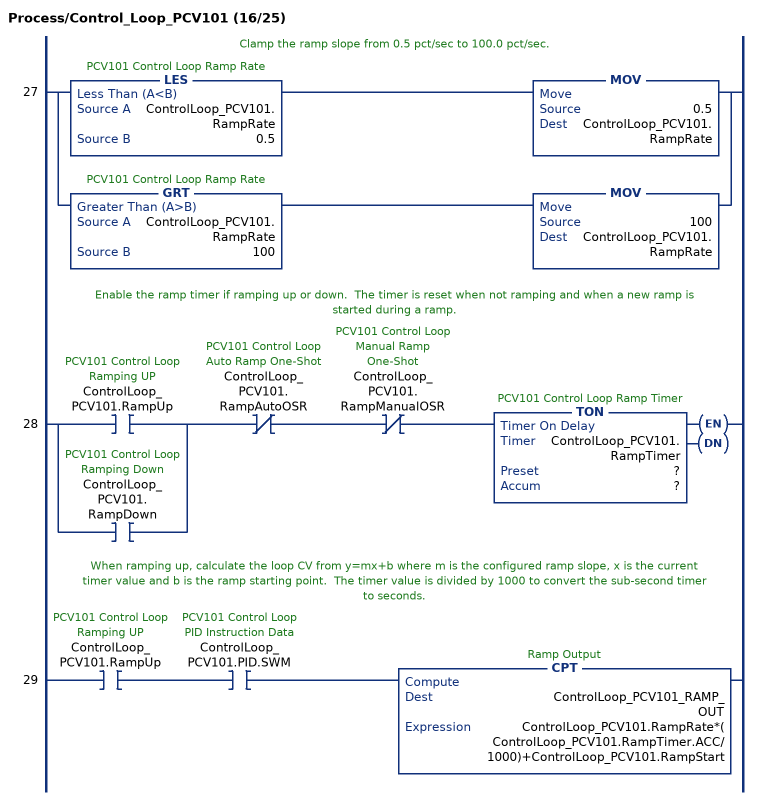
   // Clamp the ramp slope from 0.5 pct/sec to 100.0 pct/sec.
   27: [LES(ControlLoop_PCV101.RampRate,0.5) MOV(0.5,ControlLoop_PCV101.RampRate) ,GRT(ControlLoop_PCV101.RampRate,100) MOV(100,ControlLoop_PCV101.RampRate) ];
   // Enable the ramp timer if ramping up or down.  The timer is reset when not ramping and when a new ramp is started during a ramp.
   28: [XIC(ControlLoop_PCV101.RampUp) ,XIC(ControlLoop_PCV101.RampDown) ]XIO(ControlLoop_PCV101.RampAutoOSR)XIO(ControlLoop_PCV101.RampManualOSR)TON(ControlLoop_PCV101.RampTimer,?,?);
   // When ramping up, calculate the loop CV from y=mx+b where m is the configured ramp slope, x is the current timer value and b is the ramp starting point.  The timer value is divided by 1000 to convert the sub-second timer to seconds.
   29: XIC(ControlLoop_PCV101.RampUp)XIC(ControlLoop_PCV101.PID.SWM)CPT(ControlLoop_PCV101_RAMP_OUT,ControlLoop_PCV101.RampRate*(ControlLoop_PCV101.RampTimer.ACC/1000)+ControlLoop_PCV101.RampStart);
